(* IEC 61131-3 sources: avi-aoi-management/scripts/ai-eval/ngau-nhien/kho/st-ud9-ghi-dich-loai-bo/khung/src, 2 files *)

(* ---- LoaiBoAOI.st ---- *)
FUNCTION_BLOCK LoaiBoAOI
VAR_INPUT
    ENCODER : BOOL;
    CO_SAN_PHAM : BOOL;
    LOI_AOI : BOOL;
    RESET : BOOL;
    VI_TRI_GAT : INT;
    T_GAT : TIME;
END_VAR
VAR_OUTPUT
    CAN_GAT : BOOL;
    DEM_GAT : DINT;
    SO_O_LOI : INT;
END_VAR
    (* TODO: cài đặt theo đề bài *)
    CAN_GAT := FALSE;
END_FUNCTION_BLOCK

(* ---- ThanhGhiDich.st ---- *)
FUNCTION_BLOCK ThanhGhiDich
VAR_INPUT
    DICH : BOOL;
    GHI : BOOL;
    XOA : BOOL;
    VI_TRI : INT;
END_VAR
VAR_OUTPUT
    Q : BOOL;
    SO_O : INT;
END_VAR
    (* TODO: cài đặt theo đề bài *)
    Q := FALSE;
END_FUNCTION_BLOCK
